Fanuc KAREL source: KX00011.KL

PROGRAM KX00011
%NOLOCKGROUP
VAR
  I: INTEGER
  J: INTEGER
  B: BOOLEAN
  F: FILE
  S: STRING[80]
  P: XYZWPR
BEGIN
  HOLD
END KX00011
